TYPE ST_VFDError :
STRUCT
	error 	: BOOL;
	message : T_MaxString;
	
	// List flags for specific errors
	
END_STRUCT
END_TYPE

(* stored: Version 1.1.0.1, ProductVersion 3.1.4024.12
   DUT ST_VFDError: Id {6b16458b-9283-45fd-95c5-338dd23f40db} *)
